// TIA Portal V17 export
// export: Created 2026-10-28T03:24:27.1384476Z, ExportSetting WithDefaults, DisplayName Totally Integrated Automation Portal, DisplayVersion V17, DisplayName TIA Portal Openness, DisplayVersion V17, DisplayName TIA Portal Version Control Interface, DisplayVersion V17, DisplayName STEP 7 Professional, DisplayVersion V17, DisplayName STEP 7 Safety, DisplayVersion V17, DisplayName WinCC Advanced, DisplayVersion V17
TagTable "默认变量表"
  开 : Bool  (PLC tag 开, HMI_连接_1, 100 ms)
  关 : Bool  (PLC tag 关, HMI_连接_1, 100 ms)
  绿灯 : Bool  (PLC tag 绿灯, HMI_连接_1, 100 ms)
  黄灯 : Bool  (PLC tag 黄灯, HMI_连接_1, 100 ms)
  蓝灯 : Bool  (PLC tag 蓝灯, HMI_连接_1, 100 ms)
  紫灯 : Bool  (PLC tag 紫灯, HMI_连接_1, 100 ms)
  红灯 : Bool  (PLC tag 红灯, HMI_连接_1, 100 ms)
